// TIA Portal V20 export
// export: Created 2026-10-20T18:55:24.0076634Z, ExportSetting None, DisplayName Totally Integrated Automation Portal, DisplayVersion V20 Update 6, DisplayName TIA Portal Openness, DisplayVersion V20 Update 6, DisplayName TIA Portal Version Control Interface, DisplayVersion V20 Update 6, DisplayName SINAMICS Startdrive Advanced, DisplayVersion V20 SP1, DisplayName SINAMICS Startdrive G130, G150, S120, S150, SINAMICS MV, G220, S200, S210, DisplayVersion V20 SP1, DisplayName SINAMICS Startdrive G110M, G120, G120C, G120D, G120P, G115D, DisplayVersion V20 SP1, DisplayName STEP 7 Professional, DisplayVersion V20 Update 6, DisplayName STEP 7 Safety, DisplayVersion V20 Update 2, DisplayName WinCC Basic/Comfort/Advanced, DisplayVersion V20 Update 6, DisplayName WinCC Unified, DisplayVersion V20 Update 6
VAR_GLOBAL   // PLC tag table "IO_ET200_5"
   "C5105 - SENSOR CNV RIGHT (PALLET DETECT 1)" AT %I1468.4 : Bool;
   "C5107 - SENSOR CNV RIGHT (PALLET DETECT 1)" AT %I1472.4 : Bool;
   "C5103 - SENSOR CNV RIGHT (PALLET DETECT 1)" AT %I1464.4 : Bool;
   "C5104 - SENSOR CNV RIGHT (PALLET DETECT 1)" AT %I1466.4 : Bool;
   "C5101 - SENSOR CNV RIGHT (PALLET DETECT 1)" AT %I1460.4 : Bool;
   "C5108 - SENSOR CNV RIGHT (PALLET DETECT 1)" AT %I1474.4 : Bool;
   "C5102 - SENSOR CNV RIGHT (PALLET DETECT 1)" AT %I1462.4 : Bool;
   "C5106 - SENSOR CNV RIGHT (PALLET DETECT 1)" AT %I1470.4 : Bool;
   "KEY REMOTE/LOCAL L8 - CH2(5)" AT %I1750.7 : Bool;
   "E-STOP L1 - CH1(5)" AT %I1726.0 : Bool;
   "KEY REMOTE/LOCAL L1 - CH1(5)" AT %I1726.1 : Bool;
   "E-STOP L2 - CH1(5)" AT %I1726.2 : Bool;
   "KEY REMOTE/LOCAL L2 - CH1(5)" AT %I1726.3 : Bool;
   "E-STOP L1 - CH2(5)" AT %I1726.4 : Bool;
   "KEY REMOTE/LOCAL L1 - CH2(5)" AT %I1726.5 : Bool;
   "E-STOP L2 - CH2(5)" AT %I1726.6 : Bool;
   "KEY REMOTE/LOCAL L2 - CH2(5)" AT %I1726.7 : Bool;
   "E-STOP L3 - CH1(5)" AT %I1734.0 : Bool;
   "KEY REMOTE/LOCAL L3 - CH1(5)" AT %I1734.1 : Bool;
   "E-STOP L4 - CH1(5)" AT %I1734.2 : Bool;
   "KEY REMOTE/LOCAL L4 - CH1(5)" AT %I1734.3 : Bool;
   "E-STOP L3 - CH2(5)" AT %I1734.4 : Bool;
   "KEY REMOTE/LOCAL L3 - CH2(5)" AT %I1734.5 : Bool;
   "E-STOP L4 - CH2(5)" AT %I1734.6 : Bool;
   "KEY REMOTE/LOCAL L4 - CH2(5)" AT %I1734.7 : Bool;
   "E-STOP L5 - CH1(5)" AT %I1742.0 : Bool;
   "KEY REMOTE/LOCAL L5 - CH1(5)" AT %I1742.1 : Bool;
   "E-STOP L6 - CH1(5)" AT %I1742.2 : Bool;
   "KEY REMOTE/LOCAL L6 - CH1(5)" AT %I1742.3 : Bool;
   "E-STOP L5 - CH2(5)" AT %I1742.4 : Bool;
   "KEY REMOTE/LOCAL L5 - CH2(5)" AT %I1742.5 : Bool;
   "E-STOP L6 - CH2(5)" AT %I1742.6 : Bool;
   "KEY REMOTE/LOCAL L6 - CH2(5)" AT %I1742.7 : Bool;
   "E-STOP L7 - CH1(5)" AT %I1750.0 : Bool;
   "KEY REMOTE/LOCAL L7 - CH1(5)" AT %I1750.1 : Bool;
   "E-STOP L8 - CH1(5)" AT %I1750.2 : Bool;
   "KEY REMOTE/LOCAL L8 - CH1(5)" AT %I1750.3 : Bool;
   "E-STOP L7 - CH2(5)" AT %I1750.4 : Bool;
   "KEY REMOTE/LOCAL L7 - CH2(5)" AT %I1750.5 : Bool;
   "E-STOP L8 - CH2(5)" AT %I1750.6 : Bool;
   "VTD5 DOCKING PINS 1 RETRACTED" AT %I284.3 : Bool;
   "VTD5 ULTIMATE CREEP" AT %I284.5 : Bool;
   "VTD5 DOCKING PINS 2 EXTENDED" AT %I284.0 : Bool;
   "VTD5 DOCKING PINS 2 RETRACTED" AT %I284.2 : Bool;
   "VTD5 LEVEL DETECT 2" AT %I284.7 : Bool;
   "VTD5 LEVEL DETECT 1" AT %I284.6 : Bool;
   "VTD5 DOCKING PINS 1 EXTENDED" AT %I284.1 : Bool;
   "VTD5 ULTIMATE SLOWDOWN" AT %I284.4 : Bool;
   "C5102 - SENSOR SAFETY PIN1 UP" AT %I1463.2 : Bool;
   "C5101 - SHUTTLE IN POSITION 1" AT %I1461.6 : Bool;
   "C5101 - SENSOR SAFETY PIN1 UP" AT %I1461.2 : Bool;
   "C5101 - SENSOR CNV RIGHT (PALLET DETECT 2)" AT %I1461.1 : Bool;
   "C5101 - SENSOR SAFETY PIN1 DOWN" AT %I1461.3 : Bool;
   "CVTD5 SENSOR CONVEYOR CENTER" AT %I283.1 : Bool;
   "C5102 - SENSOR SAFETY PIN1 DOWN" AT %I1463.3 : Bool;
   "CVTD5 SENSOR CONVEYOR RIGHT (PALLET DETECT 1)" AT %I283.5 : Bool;
   "C5101 - SENSOR CNV LEFT (PALLET DETECT 2)" AT %I1461.0 : Bool;
   "C5101 - SENSOR CNV LEFT (FWD)" AT %I1461.4 : Bool;
   "C5101 - SENSOR CNV LEFT (PALLET DETECT 1)" AT %I1461.5 : Bool;
   "CVTD5 SENSOR CONVEYOR LEFT (PALLET DETECT 1)" AT %I283.3 : Bool;
   "CVTD5 SENSOR CONVEYOR RIGHT (BWD)" AT %I283.4 : Bool;
   "CVTD5 SENSOR CONVEYOR LEFT (FWD)" AT %I283.2 : Bool;
   "C5101 - SHUTTLE IN POSITION 2" AT %I1461.7 : Bool;
   "C5101 - SENSOR CNV RIGHT (BWD)" AT %I1460.5 : Bool;
   "C5102 - SHUTTLE IN POSITION 1" AT %I1463.6 : Bool;
   "C5102 - SENSOR CNV LEFT (PALLET DETECT 1)" AT %I1463.5 : Bool;
   "C5102 - SENSOR CNV LEFT (PALLET DETECT 2)" AT %I1463.0 : Bool;
   "C5106 - SENSOR SAFETY PIN1 DOWN" AT %I1471.3 : Bool;
   "C5108 - SENSOR SAFETY PIN1 UP" AT %I1475.2 : Bool;
   "C5107 - SENSOR CNV LEFT (FWD)" AT %I1473.4 : Bool;
   "C5107 - SENSOR CNV LEFT (PALLET DETECT 1)" AT %I1473.5 : Bool;
   "C5107 - SHUTTLE IN POSITION 1" AT %I1473.6 : Bool;
   "C5107 - SHUTTLE IN POSITION 2" AT %I1473.7 : Bool;
   "C5106 - SENSOR SAFETY PIN1 UP" AT %I1471.2 : Bool;
   "C5107 - SENSOR SAFETY PIN1 UP" AT %I1473.2 : Bool;
   "C5107 - SENSOR SAFETY PIN1 DOWN" AT %I1473.3 : Bool;
   "C5108 - SHUTTLE IN POSITION 2" AT %I1475.7 : Bool;
   "C5108 - SENSOR CNV LEFT (FWD)" AT %I1475.4 : Bool;
   "C5107 - SENSOR CNV RIGHT (PALLET DETECT 2)" AT %I1473.1 : Bool;
   "C5102 - SHUTTLE IN POSITION 2" AT %I1463.7 : Bool;
   "C5106 - SENSOR CNV LEFT (FWD)" AT %I1471.4 : Bool;
   "C5108 - SENSOR CNV LEFT (PALLET DETECT 2)" AT %I1475.0 : Bool;
   "C5107 - SENSOR CNV LEFT (PALLET DETECT 2)" AT %I1473.0 : Bool;
   "C5106 - SENSOR CNV RIGHT (PALLET DETECT 2)" AT %I1471.1 : Bool;
   "C5106 - SENSOR CNV LEFT (PALLET DETECT 2)" AT %I1471.0 : Bool;
   "C5106 - SHUTTLE IN POSITION 2" AT %I1471.7 : Bool;
   "C5106 - SENSOR CNV RIGHT (BWD)" AT %I1470.5 : Bool;
   "C5108 - SENSOR CNV RIGHT (BWD)" AT %I1474.5 : Bool;
   "C5102 - SENSOR CNV RIGHT (BWD)" AT %I1462.5 : Bool;
   "C5102 - SENSOR CNV RIGHT (PALLET DETECT 2)" AT %I1463.1 : Bool;
   "C5102 - SENSOR CNV LEFT (FWD)" AT %I1463.4 : Bool;
   "C5108 - SENSOR CNV RIGHT (PALLET DETECT 2)" AT %I1475.1 : Bool;
   "C5108 - SENSOR SAFETY PIN1 DOWN" AT %I1475.3 : Bool;
   "C5106 - SENSOR CNV LEFT (PALLET DETECT 1)" AT %I1471.5 : Bool;
   "C5108 - SENSOR CNV LEFT (PALLET DETECT 1)" AT %I1475.5 : Bool;
   "C5108 - SHUTTLE IN POSITION 1" AT %I1475.6 : Bool;
   "C5106 - SHUTTLE IN POSITION 1" AT %I1471.6 : Bool;
   "C5107 - SENSOR CNV RIGHT (BWD)" AT %I1472.5 : Bool;
   "C5105 - SENSOR CNV LEFT (FWD)" AT %I1469.4 : Bool;
   "C5105 - SENSOR SAFETY PIN1 UP" AT %I1469.2 : Bool;
   "C5103 - SENSOR CNV LEFT (PALLET DETECT 1)" AT %I1465.5 : Bool;
   "C5104 - SENSOR CNV RIGHT (PALLET DETECT 2)" AT %I1467.1 : Bool;
   "C5103 - SHUTTLE IN POSITION 1" AT %I1465.6 : Bool;
   "C5103 - SENSOR SAFETY PIN1 DOWN" AT %I1465.3 : Bool;
   "C5105 - SENSOR CNV RIGHT (BWD)" AT %I1468.5 : Bool;
   "C5104 - SENSOR CNV LEFT (PALLET DETECT 1)" AT %I1467.5 : Bool;
   "C5105 - SHUTTLE IN POSITION 2" AT %I1469.7 : Bool;
   "C5104 - SENSOR CNV LEFT (FWD)" AT %I1467.4 : Bool;
   "C5105 - SENSOR CNV LEFT (PALLET DETECT 2)" AT %I1469.0 : Bool;
   "C5103 - SENSOR CNV LEFT (PALLET DETECT 2)" AT %I1465.0 : Bool;
   "C5103 - SENSOR CNV LEFT (FWD)" AT %I1465.4 : Bool;
   "C5103 - SHUTTLE IN POSITION 2" AT %I1465.7 : Bool;
   "C5103 - SENSOR CNV RIGHT (PALLET DETECT 2)" AT %I1465.1 : Bool;
   "C5105 - SENSOR CNV RIGHT (PALLET DETECT 2)" AT %I1469.1 : Bool;
   "C5103 - SENSOR SAFETY PIN1 UP" AT %I1465.2 : Bool;
   "C5104 - SENSOR SAFETY PIN1 DOWN" AT %I1467.3 : Bool;
   "C5103 - SENSOR CNV RIGHT (BWD)" AT %I1464.5 : Bool;
   "C5105 - SENSOR CNV LEFT (PALLET DETECT 1)" AT %I1469.5 : Bool;
   "C5104 - SENSOR CNV RIGHT (BWD)" AT %I1466.5 : Bool;
   "C5104 - SENSOR SAFETY PIN1 UP" AT %I1467.2 : Bool;
   "C5104 - SENSOR CNV LEFT (PALLET DETECT 2)" AT %I1467.0 : Bool;
   "C5105 - SENSOR SAFETY PIN1 DOWN" AT %I1469.3 : Bool;
   "C5104 - SHUTTLE IN POSITION 1" AT %I1467.6 : Bool;
   "C5104 - SHUTTLE IN POSITION 2" AT %I1467.7 : Bool;
   "C5105 - SHUTTLE IN POSITION 1" AT %I1469.6 : Bool;
   "CVTD5 OVERHANG LEFT" AT %I283.7 : Bool;
   "CVTD5 OVERHANG RIGHT" AT %I283.6 : Bool;
END_VAR
